// TIA Portal V20 export
// export: Created 2026-10-19T18:04:45.0977017Z, ExportSetting WithDefaults, DisplayName Totally Integrated Automation Portal, DisplayVersion V20 Update 6, DisplayName TIA Portal Openness, DisplayVersion V20 Update 6, DisplayName TIA Portal Version Control Interface, DisplayVersion V20 Update 6, DisplayName SINAMICS Startdrive Advanced, DisplayVersion V20 SP1, DisplayName SINAMICS Startdrive G130, G150, S120, S150, SINAMICS MV, G220, S200, S210, DisplayVersion V20 SP1, DisplayName SINAMICS Startdrive G110M, G120, G120C, G120D, G120P, G115D, DisplayVersion V20 SP1, DisplayName STEP 7 Professional, DisplayVersion V20 Update 6, DisplayName STEP 7 Safety, DisplayVersion V20 Update 2, DisplayName WinCC Basic/Comfort/Advanced, DisplayVersion V20 Update 6, DisplayName WinCC Unified, DisplayVersion V20 Update 6
DATA_BLOCK "HMI_Systems"   // DB137
{ S7_Optimized_Access := 'TRUE' }
VERSION : 0.1
// stored: AutoNumber true, DBAccessibleFromOPCUA true, DBAccessibleFromWebserver true, IsOnlyStoredInLoadMemory false, IsRetainMemResEnabled false, IsWriteProtectedInAS false, MemoryReserve 100
   VAR
      SystemNo : USInt := 1;   // System Number (1 or 2)
      System { ExternalWritable := 'False'} : "System_UDT";
      CarMeasurement { ExternalWritable := 'False'} : "CarMeasurement_DB_UDT";
      EntryGate : Struct
         Sts_Opened : Bool := TRUE;
         Sts_Closed : Bool := FALSE;
         Cmd_Open : Bool := FALSE;
         Cmd_Close : Bool := FALSE;
      END_STRUCT;
      ExitGate : Struct
         Sts_Opened : Bool := TRUE;
         Sts_Closed : Bool := FALSE;
         Cmd_Open : Bool := FALSE;
         Cmd_Close : Bool := FALSE;
      END_STRUCT;
      FieldSensors : DWord := 16#04A3_7FF3;   // Field Values of Sensors
      PanelSensors : DWord := 16#04A3_7FF3;   // Sensors to show on HMI screen
      Motors : DWord := 16#0E00_6001;   // Motors to show on HMI screen
      HMI_E_Stop_System_1 : Bool := FALSE;   // HMI Emergancy Stop Push Button for System #1
      HMI_E_Stop_System_2 : Bool := FALSE;   // HMI Emergancy Stop Push Button for System #2
      HMI_E_Stop_System_3 : Bool := FALSE;   // HMI Emergancy Stop Push Button for System #2
      Virtual_Emergency_BT : Bool := false;   // HMI Emergency Stop Push Button for General system
   END_VAR
BEGIN
   System.CancelOrders := FALSE;
   System.PauseOrders := FALSE;
   System.ResumeOrders := FALSE;
   System.OrderSent := FALSE;
   System.CurrentOrder := 0;
   System.NextOrder := 1;
   System.OrderTable[0].OrderNo := 0;
   System.OrderTable[1..34].OrderNo := -1;
   System.OrderTable[35].OrderNo := 55;
   System.OrderTable[36].OrderNo := 54;
   System.OrderTable[37..38].OrderNo := 53;
   System.OrderTable[39..45].OrderNo := -1;
   System.OrderTable[46..47].OrderNo := 52;
   System.OrderTable[48..49].OrderNo := 51;
   System.OrderTable[50].OrderNo := -1;
   System.OrderTable[51].OrderNo := 50;
   System.OrderTable[52].OrderNo := 49;
   System.OrderTable[53..54].OrderNo := 48;
   System.OrderTable[55..56].OrderNo := 47;
   System.OrderTable[57..58].OrderNo := 46;
   System.OrderTable[59..60].OrderNo := 45;
   System.OrderTable[61..67].OrderNo := 44;
   System.OrderTable[68..72].OrderNo := 43;
   System.OrderTable[73..78].OrderNo := 42;
   System.OrderTable[79..80].OrderNo := 41;
   System.OrderTable[81..82].OrderNo := 40;
   System.OrderTable[83..89].OrderNo := 39;
   System.OrderTable[90..91].OrderNo := 38;
   System.OrderTable[92..96].OrderNo := 37;
   System.OrderTable[97..99].OrderNo := 36;
   System.OrderTable[0].StepNo := 0;
   System.OrderTable[1..34].StepNo := -1;
   System.OrderTable[35..36].StepNo := 1;
   System.OrderTable[37].StepNo := 2;
   System.OrderTable[38].StepNo := 1;
   System.OrderTable[39..45].StepNo := -1;
   System.OrderTable[46].StepNo := 2;
   System.OrderTable[47].StepNo := 1;
   System.OrderTable[48].StepNo := 2;
   System.OrderTable[49].StepNo := 1;
   System.OrderTable[50].StepNo := -1;
   System.OrderTable[51..52].StepNo := 1;
   System.OrderTable[53].StepNo := 2;
   System.OrderTable[54].StepNo := 1;
   System.OrderTable[55].StepNo := 2;
   System.OrderTable[56].StepNo := 1;
   System.OrderTable[57].StepNo := 2;
   System.OrderTable[58].StepNo := 1;
   System.OrderTable[59].StepNo := 2;
   System.OrderTable[60].StepNo := 1;
   System.OrderTable[61].StepNo := 7;
   System.OrderTable[62].StepNo := 6;
   System.OrderTable[63].StepNo := 5;
   System.OrderTable[64].StepNo := 4;
   System.OrderTable[65].StepNo := 3;
   System.OrderTable[66].StepNo := 2;
   System.OrderTable[67].StepNo := 1;
   System.OrderTable[68].StepNo := 5;
   System.OrderTable[69].StepNo := 4;
   System.OrderTable[70].StepNo := 3;
   System.OrderTable[71].StepNo := 2;
   System.OrderTable[72].StepNo := 1;
   System.OrderTable[73].StepNo := 6;
   System.OrderTable[74].StepNo := 5;
   System.OrderTable[75].StepNo := 4;
   System.OrderTable[76].StepNo := 3;
   System.OrderTable[77].StepNo := 2;
   System.OrderTable[78].StepNo := 1;
   System.OrderTable[79].StepNo := 2;
   System.OrderTable[80].StepNo := 1;
   System.OrderTable[81].StepNo := 2;
   System.OrderTable[82].StepNo := 1;
   System.OrderTable[83].StepNo := 7;
   System.OrderTable[84].StepNo := 6;
   System.OrderTable[85].StepNo := 5;
   System.OrderTable[86].StepNo := 4;
   System.OrderTable[87].StepNo := 3;
   System.OrderTable[88].StepNo := 2;
   System.OrderTable[89].StepNo := 1;
   System.OrderTable[90].StepNo := 2;
   System.OrderTable[91].StepNo := 1;
   System.OrderTable[92].StepNo := 5;
   System.OrderTable[93].StepNo := 4;
   System.OrderTable[94].StepNo := 3;
   System.OrderTable[95].StepNo := 2;
   System.OrderTable[96].StepNo := 1;
   System.OrderTable[97].StepNo := 6;
   System.OrderTable[98].StepNo := 5;
   System.OrderTable[99].StepNo := 4;
   System.OrderTable[0].PlaceTime := '';
   System.OrderTable[1].PlaceTime := '06/10/2022 08:58:28';
   System.OrderTable[2].PlaceTime := '06/10/2022 08:58:01';
   System.OrderTable[3].PlaceTime := '06/10/2022 08:57:38';
   System.OrderTable[4].PlaceTime := '06/10/2022 08:56:58';
   System.OrderTable[5].PlaceTime := '06/10/2022 08:46:55';
   System.OrderTable[6].PlaceTime := '06/10/2022 08:46:40';
   System.OrderTable[7].PlaceTime := '06/10/2022 08:46:00';
   System.OrderTable[8].PlaceTime := '06/10/2022 08:45:39';
   System.OrderTable[9].PlaceTime := '06/10/2022 08:45:25';
   System.OrderTable[10].PlaceTime := '06/10/2022 08:45:12';
   System.OrderTable[11].PlaceTime := '06/10/2022 08:44:47';
   System.OrderTable[12].PlaceTime := '06/10/2022 08:44:29';
   System.OrderTable[13].PlaceTime := '06/10/2022 08:44:13';
   System.OrderTable[14].PlaceTime := '06/10/2022 08:43:18';
   System.OrderTable[15].PlaceTime := '06/10/2022 08:42:58';
   System.OrderTable[16].PlaceTime := '06/10/2022 08:41:58';
   System.OrderTable[17].PlaceTime := '06/10/2022 08:41:36';
   System.OrderTable[18].PlaceTime := '06/10/2022 08:37:44';
   System.OrderTable[19].PlaceTime := '06/10/2022 08:37:27';
   System.OrderTable[20].PlaceTime := '06/10/2022 08:37:06';
   System.OrderTable[21].PlaceTime := '06/10/2022 08:35:40';
   System.OrderTable[22].PlaceTime := '06/10/2022 08:14:06';
   System.OrderTable[23].PlaceTime := '06/10/2022 08:13:36';
   System.OrderTable[24].PlaceTime := '06/10/2022 08:09:48';
   System.OrderTable[25].PlaceTime := '06/10/2022 08:09:26';
   System.OrderTable[26].PlaceTime := '06/10/2022 08:08:29';
   System.OrderTable[27].PlaceTime := '06/10/2022 08:05:42';
   System.OrderTable[28].PlaceTime := '06/10/2022 08:04:48';
   System.OrderTable[29].PlaceTime := '06/10/2022 08:03:07';
   System.OrderTable[30].PlaceTime := '06/10/2022 08:01:46';
   System.OrderTable[31].PlaceTime := '06/10/2022 08:00:57';
   System.OrderTable[32].PlaceTime := '06/10/2022 07:54:12';
   System.OrderTable[33].PlaceTime := '06/10/2022 07:53:12';
   System.OrderTable[34].PlaceTime := '06/10/2022 07:52:34';
   System.OrderTable[35].PlaceTime := '06/09/2022 15:57:28';
   System.OrderTable[36].PlaceTime := '06/09/2022 15:54:31';
   System.OrderTable[37..38].PlaceTime := '06/09/2022 15:46:22';
   System.OrderTable[39].PlaceTime := '06/09/2022 15:44:20';
   System.OrderTable[40].PlaceTime := '06/09/2022 15:44:17';
   System.OrderTable[41].PlaceTime := '06/09/2022 15:44:09';
   System.OrderTable[42].PlaceTime := '06/09/2022 15:44:07';
   System.OrderTable[43].PlaceTime := '06/09/2022 15:42:09';
   System.OrderTable[44].PlaceTime := '06/09/2022 15:42:06';
   System.OrderTable[45].PlaceTime := '06/09/2022 15:40:52';
   System.OrderTable[46..47].PlaceTime := '06/09/2022 15:38:33';
   System.OrderTable[48..49].PlaceTime := '06/09/2022 15:37:29';
   System.OrderTable[50].PlaceTime := '06/09/2022 15:28:39';
   System.OrderTable[51].PlaceTime := '06/09/2022 15:19:41';
   System.OrderTable[52].PlaceTime := '06/09/2022 15:18:44';
   System.OrderTable[53..54].PlaceTime := '06/09/2022 15:12:55';
   System.OrderTable[55..56].PlaceTime := '06/09/2022 15:06:17';
   System.OrderTable[57..58].PlaceTime := '06/09/2022 14:58:49';
   System.OrderTable[59..60].PlaceTime := '06/09/2022 14:54:55';
   System.OrderTable[61..67].PlaceTime := '06/09/2022 14:52:23';
   System.OrderTable[68..72].PlaceTime := '06/09/2022 14:50:30';
   System.OrderTable[73..78].PlaceTime := '06/09/2022 14:49:30';
   System.OrderTable[79..80].PlaceTime := '06/09/2022 14:48:13';
   System.OrderTable[81..82].PlaceTime := '06/09/2022 14:46:58';
   System.OrderTable[83..89].PlaceTime := '06/09/2022 14:44:25';
   System.OrderTable[90..91].PlaceTime := '06/09/2022 14:37:37';
   System.OrderTable[92..96].PlaceTime := '06/09/2022 14:34:13';
   System.OrderTable[97..99].PlaceTime := '06/09/2022 14:32:56';
   System.OrderTable[0].Device := '';
   System.OrderTable[1].Device := 'TurnTable';
   System.OrderTable[2].Device := 'Dolly';
   System.OrderTable[3].Device := 'TurnTable';
   System.OrderTable[4].Device := 'Dolly';
   System.OrderTable[5..36].Device := 'Shuttle';
   System.OrderTable[37].Device := 'Dolly';
   System.OrderTable[38].Device := 'Shuttle';
   System.OrderTable[39].Device := 'Dolly';
   System.OrderTable[40].Device := 'Shuttle';
   System.OrderTable[41].Device := 'Dolly';
   System.OrderTable[42].Device := 'Shuttle';
   System.OrderTable[43].Device := 'Dolly';
   System.OrderTable[44].Device := 'Shuttle';
   System.OrderTable[45..46].Device := 'Dolly';
   System.OrderTable[47].Device := 'Shuttle';
   System.OrderTable[48].Device := 'Dolly';
   System.OrderTable[49].Device := 'Shuttle';
   System.OrderTable[50].Device := 'LoadingBay Exit';
   System.OrderTable[51..52].Device := 'Shuttle';
   System.OrderTable[53].Device := 'LoadingBay Entry';
   System.OrderTable[54].Device := 'VRC';
   System.OrderTable[55].Device := 'LoadingBay Entry';
   System.OrderTable[56].Device := 'VRC';
   System.OrderTable[57].Device := 'LoadingBay Entry';
   System.OrderTable[58].Device := 'VRC';
   System.OrderTable[59].Device := 'LoadingBay Exit';
   System.OrderTable[60..61].Device := 'VRC';
   System.OrderTable[62].Device := 'Shuttle';
   System.OrderTable[63].Device := 'Dolly';
   System.OrderTable[64].Device := 'Shuttle';
   System.OrderTable[65].Device := 'Dolly';
   System.OrderTable[66].Device := 'Shuttle';
   System.OrderTable[67].Device := 'VRC';
   System.OrderTable[68].Device := 'Shuttle';
   System.OrderTable[69].Device := 'Dolly';
   System.OrderTable[70].Device := 'TurnTable';
   System.OrderTable[71].Device := 'Shuttle';
   System.OrderTable[72].Device := 'VRC';
   System.OrderTable[73].Device := 'Dolly';
   System.OrderTable[74].Device := 'CarMeasurement';
   System.OrderTable[75].Device := 'Shuttle';
   System.OrderTable[76].Device := 'TurnTable';
   System.OrderTable[77].Device := 'Shuttle';
   System.OrderTable[78].Device := 'VRC';
   System.OrderTable[79].Device := 'LoadingBay Entry';
   System.OrderTable[80].Device := 'VRC';
   System.OrderTable[81].Device := 'LoadingBay Exit';
   System.OrderTable[82..83].Device := 'VRC';
   System.OrderTable[84].Device := 'Shuttle';
   System.OrderTable[85].Device := 'Dolly';
   System.OrderTable[86].Device := 'Shuttle';
   System.OrderTable[87].Device := 'Dolly';
   System.OrderTable[88].Device := 'Shuttle';
   System.OrderTable[89].Device := 'VRC';
   System.OrderTable[90].Device := 'LoadingBay Entry';
   System.OrderTable[91].Device := 'VRC';
   System.OrderTable[92].Device := 'Shuttle';
   System.OrderTable[93].Device := 'Dolly';
   System.OrderTable[94].Device := 'TurnTable';
   System.OrderTable[95].Device := 'Shuttle';
   System.OrderTable[96].Device := 'VRC';
   System.OrderTable[97].Device := 'Dolly';
   System.OrderTable[98].Device := 'CarMeasurement';
   System.OrderTable[99].Device := 'Shuttle';
   System.OrderTable[0].Sequence := 0;
   System.OrderTable[1..61].Sequence := 1;
   System.OrderTable[62].Sequence := 0;
   System.OrderTable[63..66].Sequence := 1;
   System.OrderTable[67].Sequence := 0;
   System.OrderTable[68..71].Sequence := 1;
   System.OrderTable[72].Sequence := 0;
   System.OrderTable[73].Sequence := 1;
   System.OrderTable[74].Sequence := 0;
   System.OrderTable[75..77].Sequence := 1;
   System.OrderTable[78].Sequence := 0;
   System.OrderTable[79..83].Sequence := 1;
   System.OrderTable[84].Sequence := 0;
   System.OrderTable[85..88].Sequence := 1;
   System.OrderTable[89].Sequence := 0;
   System.OrderTable[90..95].Sequence := 1;
   System.OrderTable[96].Sequence := 0;
   System.OrderTable[97].Sequence := 1;
   System.OrderTable[98].Sequence := 0;
   System.OrderTable[99].Sequence := 1;
   System.OrderTable[0].Status := 'Error';
   System.OrderTable[1].Status := 'Completed';
   System.OrderTable[2].Status := 'Error\Cancel';
   System.OrderTable[3].Status := 'Completed';
   System.OrderTable[4].Status := 'Error\Cancel';
   System.OrderTable[5..6].Status := 'Completed';
   System.OrderTable[7].Status := 'Canceled';
   System.OrderTable[8..10].Status := 'Completed';
   System.OrderTable[11].Status := 'Canceled';
   System.OrderTable[12..15].Status := 'Completed';
   System.OrderTable[16].Status := 'Canceled';
   System.OrderTable[17..26].Status := 'Completed';
   System.OrderTable[27].Status := 'Error\Cancel';
   System.OrderTable[28..34].Status := 'Canceled';
   System.OrderTable[35..36].Status := 'Completed';
   System.OrderTable[37].Status := 'Error\Cancel';
   System.OrderTable[38..52].Status := 'Completed';
   System.OrderTable[53].Status := 'Car Refused';
   System.OrderTable[54].Status := 'Completed';
   System.OrderTable[55].Status := 'Car Refused';
   System.OrderTable[56].Status := 'Completed';
   System.OrderTable[57].Status := 'Car Refused';
   System.OrderTable[58..89].Status := 'Completed';
   System.OrderTable[90].Status := 'Car Refused';
   System.OrderTable[91..99].Status := 'Completed';
   System.OrderTable[0].CompleteTime := '06/10/2022 08:58:15';
   System.OrderTable[1].CompleteTime := '06/10/2022 08:58:44';
   System.OrderTable[2].CompleteTime := '06/10/2022 08:58:07';
   System.OrderTable[3].CompleteTime := '06/10/2022 08:57:53';
   System.OrderTable[4].CompleteTime := '06/10/2022 08:57:03';
   System.OrderTable[5].CompleteTime := '06/10/2022 08:47:08';
   System.OrderTable[6].CompleteTime := '06/10/2022 08:46:55';
   System.OrderTable[7].CompleteTime := '06/10/2022 08:46:14';
   System.OrderTable[8].CompleteTime := '06/10/2022 08:45:52';
   System.OrderTable[9].CompleteTime := '06/10/2022 08:45:38';
   System.OrderTable[10].CompleteTime := '06/10/2022 08:45:24';
   System.OrderTable[11].CompleteTime := '06/10/2022 08:44:59';
   System.OrderTable[12].CompleteTime := '06/10/2022 08:44:41';
   System.OrderTable[13].CompleteTime := '06/10/2022 08:44:28';
   System.OrderTable[14].CompleteTime := '06/10/2022 08:43:58';
   System.OrderTable[15].CompleteTime := '06/10/2022 08:43:13';
   System.OrderTable[16].CompleteTime := '06/10/2022 08:42:28';
   System.OrderTable[17].CompleteTime := '06/10/2022 08:41:49';
   System.OrderTable[18].CompleteTime := '06/10/2022 08:37:57';
   System.OrderTable[19].CompleteTime := '06/10/2022 08:37:43';
   System.OrderTable[20].CompleteTime := '06/10/2022 08:37:19';
   System.OrderTable[21].CompleteTime := '06/10/2022 08:35:45';
   System.OrderTable[22].CompleteTime := '06/10/2022 08:14:19';
   System.OrderTable[23].CompleteTime := '06/10/2022 08:13:51';
   System.OrderTable[24].CompleteTime := '06/10/2022 08:10:02';
   System.OrderTable[25].CompleteTime := '06/10/2022 08:09:37';
   System.OrderTable[26].CompleteTime := '06/10/2022 08:08:43';
   System.OrderTable[27].CompleteTime := '06/10/2022 08:07:08';
   System.OrderTable[28].CompleteTime := '06/10/2022 08:05:11';
   System.OrderTable[29].CompleteTime := '06/10/2022 08:03:33';
   System.OrderTable[30].CompleteTime := '06/10/2022 08:02:26';
   System.OrderTable[31].CompleteTime := '06/10/2022 08:01:19';
   System.OrderTable[32].CompleteTime := '06/10/2022 08:00:14';
   System.OrderTable[33].CompleteTime := '06/10/2022 07:53:22';
   System.OrderTable[34].CompleteTime := '06/10/2022 07:52:39';
   System.OrderTable[35].CompleteTime := '06/09/2022 15:57:54';
   System.OrderTable[36].CompleteTime := '06/09/2022 15:54:58';
   System.OrderTable[37].CompleteTime := '06/09/2022 15:49:19';
   System.OrderTable[38].CompleteTime := '06/09/2022 15:46:22';
   System.OrderTable[39].CompleteTime := '06/09/2022 15:45:38';
   System.OrderTable[40].CompleteTime := '06/09/2022 15:45:09';
   System.OrderTable[41].CompleteTime := '06/09/2022 15:44:52';
   System.OrderTable[42].CompleteTime := '06/09/2022 15:44:23';
   System.OrderTable[43].CompleteTime := '06/09/2022 15:42:52';
   System.OrderTable[44].CompleteTime := '06/09/2022 15:42:22';
   System.OrderTable[45].CompleteTime := '06/09/2022 15:41:22';
   System.OrderTable[46].CompleteTime := '06/09/2022 15:39:25';
   System.OrderTable[47].CompleteTime := '06/09/2022 15:38:42';
   System.OrderTable[48].CompleteTime := '06/09/2022 15:38:27';
   System.OrderTable[49].CompleteTime := '06/09/2022 15:37:44';
   System.OrderTable[50].CompleteTime := '06/09/2022 15:28:55';
   System.OrderTable[51].CompleteTime := '06/09/2022 15:19:58';
   System.OrderTable[52].CompleteTime := '06/09/2022 15:19:11';
   System.OrderTable[53].CompleteTime := '06/09/2022 15:14:08';
   System.OrderTable[54].CompleteTime := '06/09/2022 15:12:51';
   System.OrderTable[55].CompleteTime := '06/09/2022 15:07:30';
   System.OrderTable[56].CompleteTime := '06/09/2022 15:06:13';
   System.OrderTable[57].CompleteTime := '06/09/2022 15:00:22';
   System.OrderTable[58].CompleteTime := '06/09/2022 14:58:46';
   System.OrderTable[59].CompleteTime := '06/09/2022 14:56:06';
   System.OrderTable[60].CompleteTime := '06/09/2022 14:54:51';
   System.OrderTable[61].CompleteTime := '06/09/2022 14:54:47';
   System.OrderTable[62].CompleteTime := '06/09/2022 14:54:37';
   System.OrderTable[63].CompleteTime := '06/09/2022 14:54:24';
   System.OrderTable[64].CompleteTime := '06/09/2022 14:53:55';
   System.OrderTable[65].CompleteTime := '06/09/2022 14:53:33';
   System.OrderTable[66].CompleteTime := '06/09/2022 14:52:37';
   System.OrderTable[67].CompleteTime := '06/09/2022 14:52:41';
   System.OrderTable[68].CompleteTime := '06/09/2022 14:52:18';
   System.OrderTable[69].CompleteTime := '06/09/2022 14:52:00';
   System.OrderTable[70].CompleteTime := '06/09/2022 14:51:04';
   System.OrderTable[71].CompleteTime := '06/09/2022 14:50:48';
   System.OrderTable[72].CompleteTime := '06/09/2022 14:50:49';
   System.OrderTable[73].CompleteTime := '06/09/2022 14:50:25';
   System.OrderTable[74..75].CompleteTime := '06/09/2022 14:49:55';
   System.OrderTable[76].CompleteTime := '06/09/2022 14:49:43';
   System.OrderTable[77].CompleteTime := '06/09/2022 14:49:27';
   System.OrderTable[78].CompleteTime := '06/09/2022 14:49:48';
   System.OrderTable[79].CompleteTime := '06/09/2022 14:49:23';
   System.OrderTable[80].CompleteTime := '06/09/2022 14:48:10';
   System.OrderTable[81].CompleteTime := '06/09/2022 14:47:39';
   System.OrderTable[82].CompleteTime := '06/09/2022 14:46:54';
   System.OrderTable[83].CompleteTime := '06/09/2022 14:46:50';
   System.OrderTable[84].CompleteTime := '06/09/2022 14:46:41';
   System.OrderTable[85].CompleteTime := '06/09/2022 14:46:28';
   System.OrderTable[86].CompleteTime := '06/09/2022 14:45:58';
   System.OrderTable[87].CompleteTime := '06/09/2022 14:45:37';
   System.OrderTable[88].CompleteTime := '06/09/2022 14:44:40';
   System.OrderTable[89].CompleteTime := '06/09/2022 14:44:44';
   System.OrderTable[90].CompleteTime := '06/09/2022 14:38:50';
   System.OrderTable[91].CompleteTime := '06/09/2022 14:37:33';
   System.OrderTable[92].CompleteTime := '06/09/2022 14:36:02';
   System.OrderTable[93].CompleteTime := '06/09/2022 14:35:43';
   System.OrderTable[94].CompleteTime := '06/09/2022 14:34:46';
   System.OrderTable[95].CompleteTime := '06/09/2022 14:34:31';
   System.OrderTable[96].CompleteTime := '06/09/2022 14:34:32';
   System.OrderTable[97].CompleteTime := '06/09/2022 14:34:07';
   System.OrderTable[98..99].CompleteTime := '06/09/2022 14:33:36';
   System.OrderTable[0].ErrorID := 1121;
   System.OrderTable[1].ErrorID := 0;
   System.OrderTable[2].ErrorID := 1121;
   System.OrderTable[3].ErrorID := 0;
   System.OrderTable[4].ErrorID := 1117;
   System.OrderTable[5..13].ErrorID := 0;
   System.OrderTable[14].ErrorID := 2101;
   System.OrderTable[15..26].ErrorID := 0;
   System.OrderTable[27].ErrorID := 2101;
   System.OrderTable[28..31].ErrorID := 0;
   System.OrderTable[32].ErrorID := 2104;
   System.OrderTable[33..36].ErrorID := 0;
   System.OrderTable[37].ErrorID := 1118;
   System.OrderTable[38..99].ErrorID := 0;
   System.StepTable[1..20].OrderNo := 0;
   System.StepTable[1..20].StepNo := 0;
   System.StepTable[1..20].PlaceTime := '';
   System.StepTable[1..20].Device := '';
   System.StepTable[1..20].Sequence := 0;
   System.StepTable[1..20].Status := '';
   System.StepTable[1..20].CompleteTime := '';
   System.StepTable[1..20].ErrorID := 0;
   System.CarParked_Confirm := FALSE;
   System.Running := FALSE;
   System.IDLE := TRUE;
   System.Error := FALSE;
   System.State := 0;
   System.ResetError := FALSE;
   System.Ready := TRUE;
   System.Selected := TRUE;
   System.Auto_Man := TRUE;
   System.Paused := FALSE;
   CarMeasurement.Enable := TRUE;
   CarMeasurement.Execute := FALSE;
   CarMeasurement.Cancel := FALSE;
   CarMeasurement.Enabled := TRUE;
   CarMeasurement.Done := FALSE;
   CarMeasurement.Running := FALSE;
   CarMeasurement.CarSize := 0;
   CarMeasurement.strState := 'IDLE MODE';
END_DATA_BLOCK
